Fanuc KAREL source: kb00147.KL

-- PROVISIONAL review KL for V770-1; original PC SHA256 e89ce99dcaec0d0fc15b764363f75865b0e7231751979dc216c86982f9b93bce
-- Incomplete behavior may be omitted. Consult companion uncertainty JSON. Do not deploy.
PROGRAM KB00147
%NOLOCKGROUP
BEGIN
  -- UNRESOLVED_PC offsets 5-14; opcodes 3F,75
  -- UNRESOLVED_PC offsets 19-28; opcodes 3F,75
  -- UNRESOLVED_PC offsets 33-42; opcodes 3F,75
  -- UNRESOLVED_PC offsets 47-54; opcodes 9D,23
  -- UNRESOLVED_PC offsets 59-93; opcodes 27,22,2A,22,2A,22,2A,22,31
  -- UNRESOLVED_PC offsets 98-102; opcodes 7F
END KB00147
